(* IEC 61131-3 sources: codesys-framework/txt/application/WeVe Core (library)/30 Module/FB_Module, 6 files *)

(* ---- Disable.method.st ---- *)
METHOD Disable : BOOL

// --- BEGIN IMPLEMENTATION ---

IF NOT _xEnabled THEN
	Disable := TRUE;
	RETURN;
END_IF

IF _eState = E_ModuleStates.Standby THEN
	_eState := E_ModuleStates.Disable;
END_IF

(* ---- Enable.method.st ---- *)
METHOD Enable : BOOL

// --- BEGIN IMPLEMENTATION ---

IF _xEnabled THEN
	Enable := TRUE;
	RETURN;
END_IF

IF _eState = E_ModuleStates.Idle THEN
	_eState := E_ModuleStates.Enable;
END_IF

(* ---- FB_Init.method.st ---- *)
//FB_Init is always available implicitly and it is used primarily for initialization.
//The return value is not evaluated. For a specific influence, you can also declare the
//methods explicitly and provide additional code there with the standard initialization
//code. You can evaluate the return value.
METHOD FB_Init: BOOL
VAR_INPUT
    bInitRetains: BOOL; // TRUE: the retain variables are initialized (reset warm / reset cold)
    bInCopyCode: BOOL;  // TRUE: the instance will be copied to the copy code afterward (online change)

	fbEvents 	: I_EventGroup;		// de EventGroup van deze module, mag 0 zijn
END_VAR
// --- BEGIN IMPLEMENTATION ---

// Enkel de referentie bewaren, geen methodes aanroepen
_fbEvents := fbEvents;

(* ---- QuickStop.method.st ---- *)
METHOD QuickStop : BOOL

// --- BEGIN IMPLEMENTATION ---

IF _xDone THEN
	QuickStop := TRUE;
	RETURN;
END_IF

_eState := E_ModuleStates.QuickStop;

(* ---- Reset.method.st ---- *)
METHOD Reset : BOOL

// --- BEGIN IMPLEMENTATION ---

IF _xDone THEN
	Reset := TRUE;
	RETURN;
END_IF

_eState := E_ModuleStates.Reset;

(* ---- Stop.method.st ---- *)
METHOD Stop : BOOL

// --- BEGIN IMPLEMENTATION ---

IF _xDone THEN
	Stop := TRUE;
	RETURN;
END_IF

_eState := E_ModuleStates.Stop;
